Staubli VAL3: ConfProg.pjx

--- ConfProg.pjx ---
Parameters version=s7.5.3 stackSize=5000 millimeterUnit=true
Program file=MoveJoint.pgx
Program file=MoveLine.pgx
Program file=MoveCirc.pgx
Program file=start.pgx
Program file=stop.pgx
Program file=main.pgx
Data file=ConfProg.dtx

--- ConfProg.dtx ---
mdesc mNomSpeed
frame fFrame1 = {x=1234.570, y=-98.765, z=50.500, rx=-0.000, ry=0.000, rz=30.000, fatherId=world[0]}
dio Input[16]
  [0] = {link=BasicIO-1\%I0}
  [1] = {link=BasicIO-1\%I1}
  [2] = {link=BasicIO-1\%I2}
  [3] = {link=BasicIO-1\%I3}
  [4] = {link=BasicIO-1\%I4}
  [5] = {link=BasicIO-1\%I5}
  [6] = {link=BasicIO-1\%I6}
  [7] = {link=BasicIO-1\%I7}
  [8] = {link=BasicIO-1\%I8}
  [9] = {link=BasicIO-1\%I9}
  [10] = {link=BasicIO-1\%I10}
  [11] = {link=BasicIO-1\%I11}
  [12] = {link=BasicIO-1\%I12}
  [13] = {link=BasicIO-1\%I13}
  [14] = {link=BasicIO-1\%I14}
  [15] = {link=BasicIO-1\%I15}
dio Output[16]
  [0] = {link=BasicIO-1\%Q0}
  [1] = {link=BasicIO-1\%Q1}
  [2] = {link=BasicIO-1\%Q2}
  [3] = {link=BasicIO-1\%Q3}
  [4] = {link=BasicIO-1\%Q4}
  [5] = {link=BasicIO-1\%Q5}
  [6] = {link=BasicIO-1\%Q6}
  [7] = {link=BasicIO-1\%Q7}
  [8] = {link=BasicIO-1\%Q8}
  [9] = {link=BasicIO-1\%Q9}
  [10] = {link=BasicIO-1\%Q10}
  [11] = {link=BasicIO-1\%Q11}
  [12] = {link=BasicIO-1\%Q12}
  [13] = {link=BasicIO-1\%Q13}
  [14] = {link=BasicIO-1\%Q14}
  [15] = {link=BasicIO-1\%Q15}
tool tCurrentTool = {x=10.000, y=20.000, z=150.000, rx=-0.000, ry=0.000, rz=-0.000, fatherId=flange[0], ioLink=ValveIO/valve1}
mdesc mCurrentSpeed
pointRs pPointRs = {fatherId=fFrame1[0]}
pointRs pPointRs2 = {fatherId=fFrame1[0]}

--- main.pgx ---
program main()
begin
  close(tCurrentTool)
  pPointRs.config.shoulder = lefty
  pPointRs2.config.shoulder = lefty
  mCurrentSpeed.tvel = 100.00
  mCurrentSpeed.blend = joint
  mCurrentSpeed.reach = 0.010
  mCurrentSpeed.leave = 0.010
  // Program ConfProg start
  // Program generated by RoboDK v6.0.7 for Staubli TS20 FL 100 TC on XX/XX/XXXX 18:00:00
  // Using nominal kinematics.
  call MoveLine(-640.584,506.980,371.534,136.262,30.757,-130.375)
  pPointRs.config.shoulder = righty
  call MoveLine(-607.850,543.849,363.215,136.262,30.757,-130.375)
  pPointRs.config.shoulder = lefty
  call MoveLine(-602.951,596.788,316.595,136.262,30.757,-130.375)
  call MoveJoint(10.00000,20.00000,-30.00000,40.00000)
  call MoveJoint(-170.00000,45.00000,-45.00000,-170.00000)
  call MoveCirc(-353.026,-90.135,331.702,164.619,39.324,-168.579,-624.230,571.208,454.620,81.604,51.756,-128.588)

  waitEndMove()
  // Program ConfProg end

end

--- start.pgx ---
program start()
begin
  call main()
end

--- MoveCirc.pgx ---
program MoveCirc(num x_nX, num x_nY, num x_nZ, num x_nRx, num x_nRy, num x_nRz, num x_nX2, num x_nY2, num x_nZ2, num x_nRx2, num x_nRy2, num x_nRz2)
begin
  pPointRs.trsf.x = x_nX
  pPointRs.trsf.y = x_nY
  pPointRs.trsf.z = x_nZ
  pPointRs.trsf.rx = x_nRx
  pPointRs.trsf.ry = x_nRy
  pPointRs.trsf.rz = x_nRz
  pPointRs2.trsf.x = x_nX2
  pPointRs2.trsf.y = x_nY2
  pPointRs2.trsf.z = x_nZ2
  pPointRs2.trsf.rx = x_nRx2
  pPointRs2.trsf.ry = x_nRy2
  pPointRs2.trsf.rz = x_nRz2
  movec(pPointRs,pPointRs2,tCurrentTool,mCurrentSpeed)
end

--- MoveJoint.pgx ---
program MoveJoint(num x_nJ1, num x_nJ2, num x_nJ3, num x_nJ4)
  local joint l_jJoint
begin
  l_jJoint.j1 = x_nJ1
  l_jJoint.j2 = x_nJ2
  l_jJoint.j3 = x_nJ3
  l_jJoint.j4 = x_nJ4
  movej(l_jJoint,tCurrentTool ,mCurrentSpeed)
end

--- MoveLine.pgx ---
program MoveLine(num x_nX, num x_nY, num x_nZ, num x_nRx, num x_nRy, num x_nRz)
begin
  pPointRs.trsf.x = x_nX
  pPointRs.trsf.y = x_nY
  pPointRs.trsf.z = x_nZ
  pPointRs.trsf.rx = x_nRx
  pPointRs.trsf.ry = x_nRy
  pPointRs.trsf.rz = x_nRz
  movel(pPointRs,tCurrentTool,mCurrentSpeed)
end

--- stop.pgx ---
program stop()
begin
end
